TYPE ST_PTrace :		// 출력 추적표 (P, 경로 하나·그룹 하나): 위에서부터 차례로 값이 어떻게 바뀌었는지
STRUCT
	nCount		: UINT;			// 채운 줄 수
	astStep		: ARRAY[1..GVL_PARAM.TRACE_STEP_MAX] OF ST_TraceStep;
END_STRUCT
END_TYPE

(* stored: Version 1.1.0.1, ProductVersion 3.1.4024.15
   DUT ST_PTrace: Id {c3a97e12-5b4d-4f08-b6e1-92d0f8a3c574} *)
